(* IEC 61131-3 sources: sis-interlock-demo/tests/POUs/Helpers/FB_SisTestLog, 6 files *)

(* ---- CountKind.method.decl.st ---- *)
// Сколько записей кольца имеют вид eKind
METHOD CountKind : UINT
VAR_INPUT
    eKind : E_SisEventKind;   // вид события
END_VAR
VAR
    uiBack : UINT;            // сколько записей назад
    uiHits : UINT;            // найдено
    stEv   : ST_SisEvent;     // запись
END_VAR

(* ---- CountKind.method.impl.st ---- *)
uiHits := 0;
FOR uiBack := 0 TO GVL_Const.SIS_LOG_SIZE - 1 DO
    IF uiBack < uiUsed THEN
        stEv := GetEvent(uiBack := uiBack);
        IF stEv.eKind = eKind THEN
            uiHits := uiHits + 1;
        END_IF
    END_IF
END_FOR
CountKind := uiHits;

(* ---- KindAt.method.decl.st ---- *)
// Код вида записи uiBack назад (0 — последняя); вне журнала — 0 (None)
METHOD KindAt : INT
VAR_INPUT
    uiBack : UINT;            // сколько записей назад
END_VAR
VAR
    stEv : ST_SisEvent;       // запись
END_VAR

(* ---- LastOfKind.method.decl.st ---- *)
// Последняя (самая новая) запись вида eKind; нет такой — пустая запись (eKind = None)
METHOD LastOfKind : ST_SisEvent
VAR_INPUT
    eKind : E_SisEventKind;   // вид события
END_VAR
VAR
    uiBack  : UINT;           // сколько записей назад
    xFound  : BOOL;           // запись найдена
    stEv    : ST_SisEvent;    // запись
    stFound : ST_SisEvent;    // результат
END_VAR

(* ---- LastOfKind.method.impl.st ---- *)
xFound := FALSE;
FOR uiBack := 0 TO GVL_Const.SIS_LOG_SIZE - 1 DO
    IF NOT xFound AND uiBack < uiUsed THEN
        stEv := GetEvent(uiBack := uiBack);
        IF stEv.eKind = eKind THEN
            stFound := stEv;
            xFound := TRUE;
        END_IF
    END_IF
END_FOR
LastOfKind := stFound;

(* ---- SetSeq.method.decl.st ---- *)
// Установить номер последнего события (только для тестов перехода номера через 16#FFFFFFFF)
METHOD SetSeq
VAR_INPUT
    udiValue : UDINT;   // новый номер последнего события
END_VAR
